(* IEC 61131-3 sources: llm-plc-st-eval/data/definitivo/claude-sonnet-4-6/I5/zero_shot, 3 files *)

(* ---- ejec_1.st ---- *)
```pascal
FUNCTION_BLOCK FB_Clasificadora
VAR_INPUT
    sensorPresencia : BOOL; (* Sensor de paso de pieza *)
    sensorAltura    : BOOL; (* TRUE = pieza alta *)
END_VAR

VAR_OUTPUT
    banda   : BOOL; (* Salida banda transportadora *)
    piston  : BOOL; (* Salida pistón desviador *)
    nAltas  : INT;  (* Contador de piezas altas *)
    nBajas  : INT;  (* Contador de piezas bajas *)
END_VAR

VAR
    tRetardo    : TON; (* Temporizador retardo 2 s hasta el desviador *)
    tPiston     : TON; (* Temporizador duración del pistón 1 s *)
    rPresencia  : R_TRIG; (* Flanco ascendente del sensor de presencia *)
    bPiezaAlta  : BOOL;  (* Memoriza si la pieza detectada es alta *)
    bEsperando  : BOOL;  (* TRUE mientras se espera el retardo de 2 s *)
END_VAR

(* ── Banda siempre activa ─────────────────────────────────────── *)
banda := TRUE;

(* ── Detección de flanco en sensorPresencia ───────────────────── *)
rPresencia(CLK := sensorPresencia);

IF rPresencia.Q THEN
    (* Nueva pieza detectada; registrar su tipo y arrancar retardo *)
    bPiezaAlta := sensorAltura;

    IF bPiezaAlta THEN
        nAltas := nAltas + 1; (* Contar pieza alta *)
        bEsperando := TRUE;   (* Activar espera del retardo *)
    ELSE
        nBajas := nBajas + 1; (* Contar pieza baja; no se desvía *)
    END_IF;
END_IF;

(* ── Temporizador de retardo: 2 s desde detección ────────────── *)
tRetardo(IN := bEsperando, PT := T#2S);

IF tRetardo.Q THEN
    (* Han pasado 2 s: activar pistón y arrancar su temporizador *)
    bEsperando := FALSE;
    tRetardo(IN := FALSE); (* Resetear temporizador de retardo *)
END_IF;

(* ── Temporizador de duración del pistón: 1 s ────────────────── *)
tPiston(IN := tRetardo.Q, PT := T#1S);
(* Nota: tRetardo.Q permanece TRUE un ciclo; el flanco es suficiente
   para que tPiston arranque con IN=TRUE en ese ciclo.             *)

piston := tPiston.IN AND NOT tPiston.Q;
(* El pistón está activo mientras tPiston cuenta y aún no terminó *)

IF tPiston.Q THEN
    tPiston(IN := FALSE); (* Resetear temporizador del pistón *)
END_IF;

END_FUNCTION_BLOCK
```

> **Notas de diseño**
>
> | Elemento | Decisión |
> |---|---|
> | `banda` | Siempre `TRUE`; la banda nunca se detiene. |
> | `R_TRIG` | Garantiza que cada pieza se procesa una sola vez aunque el sensor permanezca activo varios ciclos. |
> | `bPiezaAlta` | Memoriza el tipo de pieza durante los 2 s de retardo. |
> | `tRetardo` (TON, `T#2S`) | Modela el tiempo de tránsito pieza → desviador. |
> | `tPiston` (TON, `T#1S`) | Controla la duración de la activación del pistón. |
> | Contadores | Se incrementan en el momento de la detección, antes de que la pieza llegue al desviador. |

(* ---- ejec_2.st ---- *)
```pascal
FUNCTION_BLOCK FB_Clasificadora
VAR_INPUT
    sensorPresencia : BOOL; (* Sensor de paso de pieza *)
    sensorAltura    : BOOL; (* TRUE = pieza alta *)
END_VAR

VAR_OUTPUT
    banda   : BOOL; (* Banda transportadora activa *)
    piston  : BOOL; (* Pistón desviador *)
    nAltas  : INT;  (* Contador de piezas altas *)
    nBajas  : INT;  (* Contador de piezas bajas *)
END_VAR

VAR
    tRetardo    : TON; (* Temporizador retardo 2 s hasta el desviador *)
    tPiston     : TON; (* Temporizador duración del pistón 1 s *)
    rPresencia  : R_TRIG; (* Flanco ascendente del sensor de presencia *)
    bPiezaAlta  : BOOL;  (* Indica que la pieza detectada es alta *)
    bContado    : BOOL;  (* Evita contar la misma pieza más de una vez *)
END_VAR

(* ------------------------------------------------------------------ *)
(* 1. La banda funciona siempre                                        *)
(* ------------------------------------------------------------------ *)
banda := TRUE;

(* ------------------------------------------------------------------ *)
(* 2. Detectar flanco ascendente del sensor de presencia              *)
(* ------------------------------------------------------------------ *)
rPresencia(CLK := sensorPresencia);

IF rPresencia.Q THEN
    (* Capturar si la pieza es alta en el momento de la detección *)
    bPiezaAlta := sensorAltura;
    bContado   := FALSE; (* Reiniciar bandera de conteo *)

    IF bPiezaAlta THEN
        (* Arrancar el temporizador de retardo (2 s) *)
        tRetardo.IN := FALSE; (* Reset previo para reiniciar *)
    END_IF;
END_IF;

(* ------------------------------------------------------------------ *)
(* 3. Temporizador de retardo: 2 s desde la detección                 *)
(* ------------------------------------------------------------------ *)
tRetardo(IN := bPiezaAlta AND NOT tPiston.Q,
         PT := T#2S);

(* ------------------------------------------------------------------ *)
(* 4. Temporizador de pistón: 1 s de activación                       *)
(* ------------------------------------------------------------------ *)
tPiston(IN := tRetardo.Q,
        PT := T#1S);

(* ------------------------------------------------------------------ *)
(* 5. Activar pistón durante el tiempo definido                       *)
(* ------------------------------------------------------------------ *)
piston := tPiston.IN AND NOT tPiston.Q;
(* tPiston.IN=TRUE y Q=FALSE => dentro del período de 1 s            *)

(* ------------------------------------------------------------------ *)
(* 6. Cuando el pistón termina, limpiar estado y contar               *)
(* ------------------------------------------------------------------ *)
IF tPiston.Q AND NOT bContado THEN
    nAltas   := nAltas + 1;
    bContado   := TRUE;
    bPiezaAlta := FALSE; (* Liberar para la siguiente pieza *)
    tRetardo.IN := FALSE; (* Reiniciar temporizadores *)
    tPiston.IN  := FALSE;
END_IF;

(* ------------------------------------------------------------------ *)
(* 7. Contar piezas bajas (flanco de presencia + altura inactiva)     *)
(* ------------------------------------------------------------------ *)
IF rPresencia.Q AND NOT sensorAltura THEN
    nBajas := nBajas + 1;
END_IF;

END_FUNCTION_BLOCK
```

(* ---- ejec_3.st ---- *)
```pascal
FUNCTION_BLOCK FB_Clasificadora
VAR_INPUT
    sensorPresencia : BOOL; (* Detecta el paso de una pieza *)
    sensorAltura    : BOOL; (* TRUE si la pieza es alta *)
END_VAR

VAR_OUTPUT
    banda   : BOOL; (* Activa la banda transportadora *)
    piston  : BOOL; (* Activa el desviador *)
    nAltas  : INT;  (* Contador de piezas altas *)
    nBajas  : INT;  (* Contador de piezas bajas *)
END_VAR

VAR
    rPresencia      : R_TRIG;       (* Flanco ascendente de sensorPresencia *)
    piezaAlta       : BOOL;         (* Indica que la pieza detectada es alta *)
    timerRetardo    : TON;          (* Retardo de 2 s hasta el desviador *)
    timerPiston     : TON;          (* Duración de 1 s del pistón *)
END_VAR

(* ─────────────────────────────────────────────
   La banda funciona siempre de forma continua
   ───────────────────────────────────────────── *)
banda := TRUE;

(* ─────────────────────────────────────────────
   Detección de flanco ascendente en sensorPresencia
   ───────────────────────────────────────────── *)
rPresencia(CLK := sensorPresencia);

IF rPresencia.Q THEN
    (* Nueva pieza detectada *)
    IF sensorAltura THEN
        (* Pieza alta: armar retardo y contabilizar *)
        piezaAlta := TRUE;
        nAltas    := nAltas + 1;
    ELSE
        (* Pieza baja: solo contabilizar *)
        nBajas := nBajas + 1;
    END_IF;
END_IF;

(* ─────────────────────────────────────────────
   Temporizador de retardo: 2 s desde la detección
   Se activa mientras piezaAlta esté pendiente y
   el pistón aún no haya comenzado su ciclo
   ───────────────────────────────────────────── *)
timerRetardo(IN := piezaAlta AND NOT timerPiston.Q,
             PT := T#2S);

(* ─────────────────────────────────────────────
   Temporizador del pistón: 1 s de activación
   Arranca cuando el retardo ha concluido
   ───────────────────────────────────────────── *)
timerPiston(IN := timerRetardo.Q,
            PT := T#1S);

(* ─────────────────────────────────────────────
   Salida del pistón activa durante el segundo
   temporizador
   ───────────────────────────────────────────── *)
piston := timerPiston.IN AND NOT timerPiston.Q;

(* ─────────────────────────────────────────────
   Cuando el pistón termina su ciclo, limpiar
   el flag y dejar que los temporizadores se
   reinicien en el siguiente ciclo de scan
   ───────────────────────────────────────────── *)
IF timerPiston.Q THEN
    piezaAlta := FALSE;
END_IF;

END_FUNCTION_BLOCK
```
